# EPICS autosave request: iocs/motor/smaract-ioc/auto_positions.req
file "asyn_motor_positions.req", P=$(P), M=m1
file "asyn_motor_positions.req", P=$(P), M=m2
file "asyn_motor_positions.req", P=$(P), M=m3
